DATA_BLOCK "naut_Tags"
{ S7_Optimized_Access := 'TRUE' }
VERSION : 0.1
   VAR
      Go : BOOL;
      N : DINT;
      Out : BOOL;
   END_VAR

BEGIN

END_DATA_BLOCK
